(* IEC 61131-3 sources: llm-plc-st-eval/data/raw/claude-sonnet-4-6/B1/few_shot, 3 files *)

(* ---- ejec_1.st ---- *)
```pascal
FUNCTION_BLOCK FB_Motor
VAR_INPUT
    btnMarcha : BOOL; (* Boton de marcha (NA) *)
    btnParo   : BOOL; (* Boton de paro (NC, activo = paro) *)
    btnEmerg  : BOOL; (* Paro de emergencia (NC, activo = emergencia) *)
END_VAR
VAR_OUTPUT
    motorOn : BOOL; (* Contactor / salida del motor *)
END_VAR
VAR
    bloqEmerg : BOOL; (* Bloqueo activo tras paro de emergencia *)
END_VAR

(* Activar bloqueo de emergencia con flanco o nivel de btnEmerg *)
IF btnEmerg THEN
    bloqEmerg := TRUE;
END_IF;

(* Reset del bloqueo: solo cuando la emergencia este liberada Y el motor este parado *)
IF NOT btnEmerg AND NOT motorOn THEN
    bloqEmerg := FALSE;
END_IF;

(* Logica de arranque/paro con autoretencion *)
(* Paro tiene prioridad sobre marcha; bloqueo impide rearranque tras emergencia *)
IF btnParo OR btnEmerg THEN
    motorOn := FALSE;                              (* Paro normal o emergencia *)
ELSIF btnMarcha AND NOT bloqEmerg THEN
    motorOn := TRUE;                               (* Arranque solo si no hay bloqueo *)
END_IF;

END_FUNCTION_BLOCK
```

(* ---- ejec_2.st ---- *)
```st
FUNCTION_BLOCK FB_Motor
VAR_INPUT
    btnMarcha : BOOL; (* Boton de marcha *)
    btnParo   : BOOL; (* Boton de paro *)
    btnEmerg  : BOOL; (* Boton de paro de emergencia *)
END_VAR
VAR_OUTPUT
    motorOn : BOOL; (* Salida del contactor del motor *)
END_VAR
VAR
    bloqEmerg : BOOL; (* Bloqueo activo tras paro de emergencia *)
END_VAR

(* Activar bloqueo ante paro de emergencia; se mantiene hasta que
   btnMarcha se suelte, evitando un rearranque involuntario *)
IF btnEmerg THEN
    bloqEmerg := TRUE;
END_IF;

(* Liberar bloqueo solo cuando el operador suelte el boton de marcha *)
IF bloqEmerg AND NOT btnMarcha THEN
    bloqEmerg := FALSE;
END_IF;

(* Logica de arranque/paro con autoretencion:
   - SET:   btnMarcha activo y sin bloqueo de emergencia
   - RESET: btnParo, btnEmerg o bloqueo activo *)
IF btnMarcha AND NOT bloqEmerg THEN
    motorOn := TRUE;
END_IF;

IF btnParo OR btnEmerg OR bloqEmerg THEN
    motorOn := FALSE;
END_IF;

END_FUNCTION_BLOCK
```

(* ---- ejec_3.st ---- *)
```pascal
FUNCTION_BLOCK FB_Motor
VAR_INPUT
    btnMarcha : BOOL; (* Boton de marcha (NA) *)
    btnParo   : BOOL; (* Boton de paro (NC, activo = paro) *)
    btnEmerg  : BOOL; (* Paro de emergencia (NC, activo = emergencia) *)
END_VAR
VAR_OUTPUT
    motorOn : BOOL; (* Contactor / salida del motor *)
END_VAR
VAR
    bloqEmerg : BOOL; (* Bloqueo activo tras paro de emergencia *)
END_VAR

(* Activar bloqueo de emergencia con flanco o nivel de btnEmerg *)
IF btnEmerg THEN
    bloqEmerg := TRUE;
END_IF;

(* Resetear bloqueo solo cuando la emergencia este liberada y el motor este parado *)
IF NOT btnEmerg AND NOT motorOn THEN
    bloqEmerg := FALSE;
END_IF;

(* Logica de arranque/paro con autoretencion:
   - Arranca : btnMarcha activo, sin paro, sin emergencia y sin bloqueo
   - Para    : btnParo o btnEmerg activos                               *)
IF (btnParo OR btnEmerg) THEN
    motorOn := FALSE;
ELSIF (btnMarcha AND NOT bloqEmerg) THEN
    motorOn := TRUE;
END_IF;

END_FUNCTION_BLOCK
```
